FUNCTION ExportFunction (* Function exported as service interface function *)
  (* Standard: 61499-1; Description: Copyright (c) 2026 Osoft e.U. This program and the accompanying materials are made available under the terms of the Eclipse Public License 2.0 which is available at https://www.eclipse.org/legal/epl-2.0/ SPDX-License-Identifier: EPL-2.0 *)
  (* Version 1.0, 2026-11-19, Michael Oberlehner, initial API and implementation and/or initial documentation *)
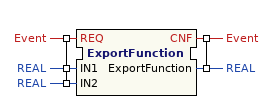
  EVENT_INPUT
    REQ WITH IN1, IN2;
  END_EVENT
  EVENT_OUTPUT
    CNF WITH ExportFunction;
  END_EVENT
  VAR_INPUT
    IN1 : REAL;
    IN2 : REAL;
  END_VAR
  VAR_OUTPUT
    ExportFunction : REAL;
  END_VAR
  BODY IN ST:
FUNCTION ExportFunction : REAL
VAR_INPUT
	IN1 : REAL;
	IN2 : REAL;
END_VAR

ExportFunction := IN1 + IN2;

END_FUNCTION
  END_BODY
END_FUNCTION
